Fanuc KAREL source: ka00215.KL

-- PROVISIONAL review KL for V1013-1; original PC SHA256 7856ea7e687f6c317fb52526084097f13e11722a571a2e0567ddc789ee98f05e
-- Incomplete behavior may be omitted. Consult companion uncertainty JSON. Do not deploy.
PROGRAM KA00215
%NOLOCKGROUP
BEGIN
  -- UNRESOLVED_PC offsets 5-19; opcodes 22,22,1E
  -- UNRESOLVED_PC offsets 24-28; opcodes 7F
END KA00215
